PROGRAM main
  VAR
    S1 AT %IX0.0  : BOOL; (* arranque *)
    B1 AT %IX0.1  : BOOL; (* presencia (selector) *)
    H1 AT %QX0.0  : BOOL; (* arranque *)
    H2 AT %QX0.1  : BOOL; (* luz del pasillo *)
    HA1 AT %QX0.2 : BOOL; (* bocina *)
    ARRANQUE      : TON;
    PASILLO       : TOF;
    BOCINA        : TON;
  END_VAR

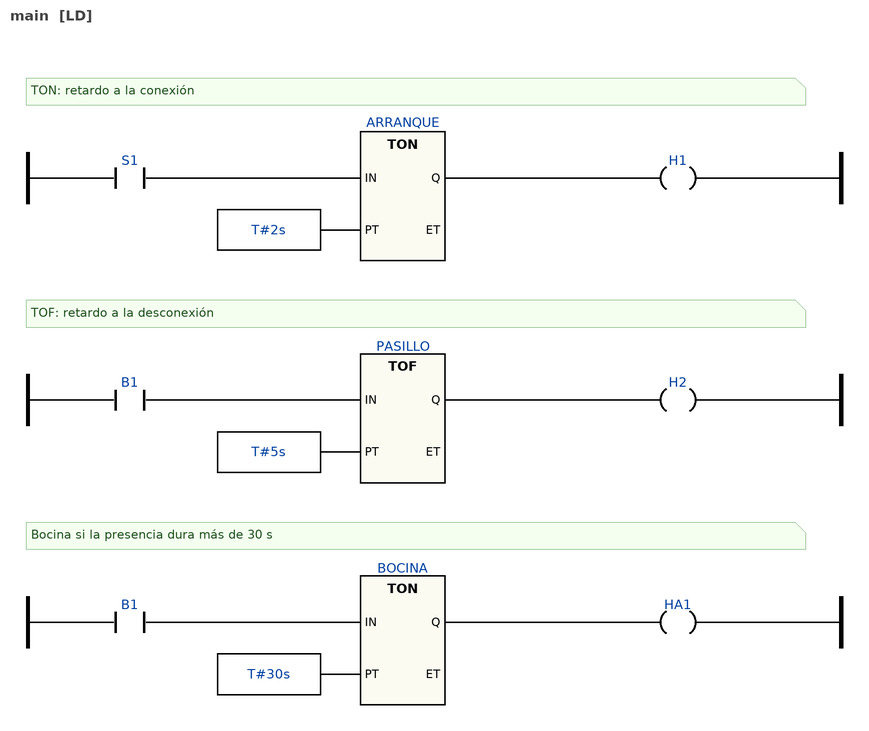
(* LD diagram, written out as Structured Text *)
(* TON: retardo a la conexión *)
ARRANQUE(IN := S1, PT := T#2s);
H1 := ARRANQUE.Q;
(* TOF: retardo a la desconexión *)
PASILLO(IN := B1, PT := T#5s);
H2 := PASILLO.Q;
(* Bocina si la presencia dura más de 30 s *)
BOCINA(IN := B1, PT := T#30s);
HA1 := BOCINA.Q;
END_PROGRAM
